// TIA Portal V20 export
// export: Created 2026-11-17T22:08:17.5244269Z, ExportSetting WithDefaults, DisplayName Totally Integrated Automation Portal, DisplayVersion V20 Update 7, DisplayName TIA Portal Openness, DisplayVersion V20 Update 7, DisplayName TIA Portal Version Control Interface, DisplayVersion V20 Update 7, DisplayName TIA Portal Test Suite Advanced, DisplayVersion V20, DisplayName SINAMICS Startdrive Advanced, DisplayVersion V20 SP1 Update 1, DisplayName SINAMICS Startdrive G110M, G120, G120C, G120D, G120P, G115D, DisplayVersion V20 SP1 Update 1, DisplayName SINAMICS Startdrive G130, G150, S120, S150, SINAMICS MV, G220, S200, S210, DisplayVersion V20 SP1 Update 1, DisplayName STEP 7 Professional, DisplayVersion V20 Update 7, DisplayName STEP 7 Safety, DisplayVersion V20 Update 2, DisplayName WinCC Basic/Comfort/Advanced, DisplayVersion V20 Update 7, DisplayName WinCC Unified, DisplayVersion V20 Update 7
FUNCTION_BLOCK "zzE2eFbd"   // FB7, FBD
{ S7_Optimized_Access := 'TRUE' }
VERSION : 0.1
// stored: AutoNumber true, IsIECCheckEnabled false, IsRetainMemResEnabled false, MemoryReserve 100, SetENOAutomatically false, UDAEnableTagReadback false
   VAR_INPUT
      ina : Bool;
      inb : Bool;
      inc : Bool;
      ind : Bool;
      iv1 : Int;
      iv2 : Int;
   END_VAR
   VAR_OUTPUT
      outq : Bool;
      outr : Bool;
      ov1 : Int;
   END_VAR
BEGIN

REGION Network 1: And gate
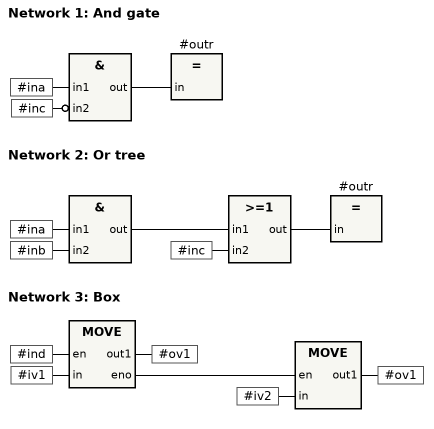
   #outr := #ina AND NOT #inc;
END_REGION

REGION Network 2: Or tree
   #outr := (#ina AND #inb) OR #inc;
END_REGION

REGION Network 3: Box
   // ENO of a box is taken as its EN; it also drops when the box reports an error
   IF #ind THEN
       #ov1 := #iv1;
       #ov1 := #iv2;
   END_IF;
END_REGION
END_FUNCTION_BLOCK
